// Mitsubishi GX Works2 project: Ex_2   PLC: FX3G

PROGRAM MAIN
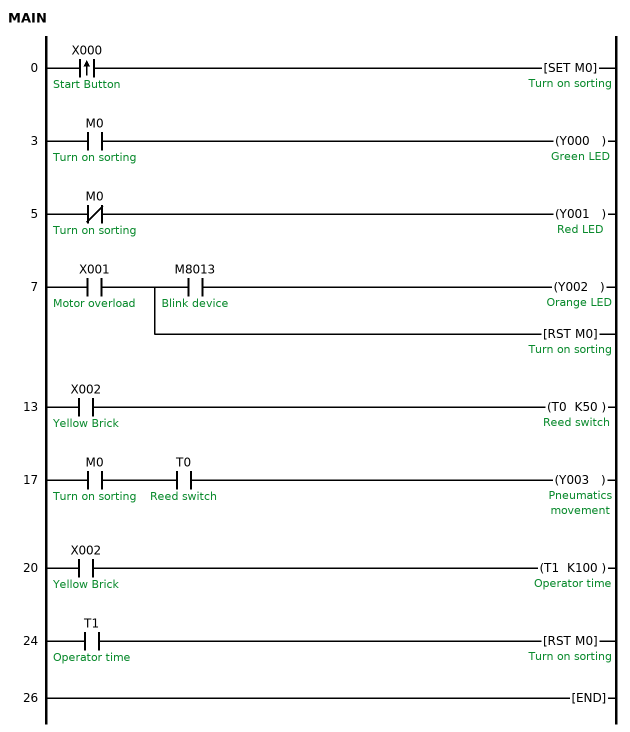
0     LDP     X000  ; Start Button
      SET     M0  ; Turn on sorting
3     LD      M0  ; Turn on sorting
      OUT     Y000  ; Green LED
5     LDI     M0  ; Turn on sorting
      OUT     Y001  ; Red LED
7     LD      X001  ; Motor overload
      MPS
      AND     M8013  ; Blink device
      OUT     Y002  ; Orange LED
      MPP
      RST     M0  ; Turn on sorting
13    LD      X002  ; Yellow Brick
      OUT     T0 K50  ; Reed switch
17    LD      M0  ; Turn on sorting
      AND     T0  ; Reed switch
      OUT     Y003  ; Pneumatics movement
20    LD      X002  ; Yellow Brick
      OUT     T1 K100  ; Operator time
24    LD      T1  ; Operator time
      RST     M0  ; Turn on sorting
26    END
END_PROGRAM
